(* IEC 61131-3 sources: avi-aoi-management/scripts/ai-eval/ngau-nhien/kho/st-ud2-den-giao-thong/mau/src, 2 files *)

(* ---- DenGiaoThong.st ---- *)
FUNCTION_BLOCK DenGiaoThong
VAR_INPUT
    NUT_NGUOI : BOOL;
    NHAP_NHAY_VANG : BOOL;
    T_XANH_MIN : TIME;
    T_VANG : TIME;
    T_NGUOI : TIME;
    T_DO_CHUNG : TIME;
    T_NHAY : TIME;
END_VAR
VAR_OUTPUT
    XE_XANH : BOOL;
    XE_VANG : BOOL;
    XE_DO : BOOL;
    NG_XANH : BOOL;
    NG_DO : BOOL;
    TRANG_THAI : INT;  (* 0 XANH_XE, 1 VANG, 2 NGUOI_DI, 3 DO_CHUNG, 4 NHAP_NHAY *)
END_VAR
VAR
    nn : NhapNhay;
    tBuoc : TON;       (* ET = thời gian đã ở trạng thái hiện tại *)
    yeuCau : BOOL;
    ttTruoc : INT;
END_VAR
    tBuoc(IN := TRUE, PT := T#24h);
    IF NUT_NGUOI AND TRANG_THAI = 0 THEN
        yeuCau := TRUE;
    END_IF

    IF NHAP_NHAY_VANG THEN
        TRANG_THAI := 4;
    ELSE
        CASE TRANG_THAI OF
        0: IF yeuCau AND tBuoc.ET >= T_XANH_MIN THEN TRANG_THAI := 1; END_IF
        1: IF tBuoc.ET >= T_VANG THEN TRANG_THAI := 2; END_IF
        2: IF tBuoc.ET >= T_NGUOI THEN TRANG_THAI := 3; END_IF
        3: IF tBuoc.ET >= T_DO_CHUNG THEN TRANG_THAI := 0; END_IF
        4: TRANG_THAI := 3;
        END_CASE
    END_IF
    IF TRANG_THAI <> 0 THEN
        yeuCau := FALSE;
    END_IF
    IF TRANG_THAI <> ttTruoc THEN
        tBuoc(IN := FALSE);
        tBuoc(IN := TRUE, PT := T#24h);
    END_IF
    ttTruoc := TRANG_THAI;

    nn(EN := TRANG_THAI = 4, T_NUA := T_NHAY);
    XE_XANH := TRANG_THAI = 0;
    XE_VANG := TRANG_THAI = 1 OR (TRANG_THAI = 4 AND nn.Q);
    XE_DO := TRANG_THAI = 2 OR TRANG_THAI = 3;
    NG_XANH := TRANG_THAI = 2;
    NG_DO := TRANG_THAI = 0 OR TRANG_THAI = 1 OR TRANG_THAI = 3;
END_FUNCTION_BLOCK

(* ---- NhapNhay.st ---- *)
FUNCTION_BLOCK NhapNhay
VAR_INPUT
    EN : BOOL;
    T_NUA : TIME;
END_VAR
VAR_OUTPUT
    Q : BOOL;
END_VAR
VAR
    tDao : TON;
    dangBat : BOOL;
END_VAR
    IF NOT EN THEN
        Q := FALSE;
        dangBat := FALSE;
        tDao(IN := FALSE);
    ELSE
        IF NOT dangBat THEN
            dangBat := TRUE;
            Q := TRUE;
            tDao(IN := FALSE);
        END_IF
        tDao(IN := TRUE, PT := T_NUA);
        IF tDao.Q THEN
            Q := NOT Q;
            tDao(IN := FALSE);
            tDao(IN := TRUE, PT := T_NUA);
        END_IF
    END_IF
END_FUNCTION_BLOCK
